(* IEC 61131-3 sources: plc-st-coding-agent/progress/evidence/f14_v2_public_20261112b/jobs/codex_minimax-m27, 5 files *)

(* ---- public-easy-01.candidate_01.st ---- *)
FUNCTION_BLOCK FillingLineControl
VAR_INPUT
    bottleSensor           : BOOL;
    cleaningConfirmButton  : BOOL;
    fillingConfirmButton   : BOOL;
    cappingConfirmButton   : BOOL;
    packingConfirmButton   : BOOL;
    finishedButton         : BOOL;
END_VAR

VAR_OUTPUT
    Pump_Motor     : BOOL := FALSE;
    Filling_Valve  : BOOL := FALSE;
    Capping_Machine: BOOL := FALSE;
    Packing_Machine: BOOL := FALSE;
    Completion_Light: BOOL := FALSE;
END_VAR

VAR
    state : INT := 0;
    lastBottleSensor : BOOL := FALSE;
END_VAR

    // Detect bottle arrival
    IF bottleSensor AND NOT lastBottleSensor THEN
        state := 1;
    END_IF
    lastBottleSensor := bottleSensor;

    // State machine
    CASE state OF
        0:  // IDLE
            Pump_Motor := FALSE;
            Filling_Valve := FALSE;
            Capping_Machine := FALSE;
            Packing_Machine := FALSE;
            Completion_Light := FALSE;

        1:  // CLEANING
            Pump_Motor := TRUE;
            Filling_Valve := FALSE;
            Capping_Machine := FALSE;
            Packing_Machine := FALSE;
            Completion_Light := FALSE;
            IF cleaningConfirmButton THEN
                state := 2;
            END_IF

        2:  // FILLING
            Pump_Motor := FALSE;
            Filling_Valve := TRUE;
            Capping_Machine := FALSE;
            Packing_Machine := FALSE;
            Completion_Light := FALSE;
            IF fillingConfirmButton THEN
                state := 3;
            END_IF

        3:  // CAPPING
            Pump_Motor := FALSE;
            Filling_Valve := FALSE;
            Capping_Machine := TRUE;
            Packing_Machine := FALSE;
            Completion_Light := FALSE;
            IF cappingConfirmButton THEN
                state := 4;
            END_IF

        4:  // PACKING
            Pump_Motor := FALSE;
            Filling_Valve := FALSE;
            Capping_Machine := FALSE;
            Packing_Machine := TRUE;
            Completion_Light := FALSE;
            IF packingConfirmButton THEN
                state := 5;
            END_IF

        5:  // COMPLETE
            Pump_Motor := FALSE;
            Filling_Valve := FALSE;
            Capping_Machine := FALSE;
            Packing_Machine := FALSE;
            Completion_Light := TRUE;
            IF finishedButton THEN
                state := 0;
            END_IF
    END_CASE
END_FUNCTION_BLOCK

(* ---- public-easy-01.candidate_02.st ---- *)
FUNCTION_BLOCK FillingLineControl
VAR_INPUT
    bottleSensor           : BOOL;
    cleaningConfirmButton  : BOOL;
    fillingConfirmButton   : BOOL;
    cappingConfirmButton   : BOOL;
    packingConfirmButton   : BOOL;
    finishedButton         : BOOL;
END_VAR

VAR_OUTPUT
    Pump_Motor      : BOOL := FALSE;
    Filling_Valve   : BOOL := FALSE;
    Capping_Machine : BOOL := FALSE;
    Packing_Machine : BOOL := FALSE;
    Completion_Light: BOOL := FALSE;
END_VAR

VAR
    state               : INT := 0;
    lastBottleSensor    : BOOL := FALSE;
    lastCleaningButton  : BOOL := FALSE;
    lastFillingButton   : BOOL := FALSE;
    lastCappingButton   : BOOL := FALSE;
    lastPackingButton   : BOOL := FALSE;
    lastFinishedButton  : BOOL := FALSE;
END_VAR

    // Detect bottle arrival on rising edge
    IF bottleSensor AND NOT lastBottleSensor THEN
        state := 1;
    END_IF
    lastBottleSensor := bottleSensor;

    // State machine
    CASE state OF
        0:  // IDLE
            Pump_Motor := FALSE;
            Filling_Valve := FALSE;
            Capping_Machine := FALSE;
            Packing_Machine := FALSE;
            Completion_Light := FALSE;

        1:  // CLEANING
            Pump_Motor := TRUE;
            Filling_Valve := FALSE;
            Capping_Machine := FALSE;
            Packing_Machine := FALSE;
            Completion_Light := FALSE;
            // Rising edge detection for button
            IF cleaningConfirmButton AND NOT lastCleaningButton THEN
                state := 2;
            END_IF

        2:  // FILLING
            Pump_Motor := FALSE;
            Filling_Valve := TRUE;
            Capping_Machine := FALSE;
            Packing_Machine := FALSE;
            Completion_Light := FALSE;
            // Rising edge detection for button
            IF fillingConfirmButton AND NOT lastFillingButton THEN
                state := 3;
            END_IF

        3:  // CAPPING
            Pump_Motor := FALSE;
            Filling_Valve := FALSE;
            Capping_Machine := TRUE;
            Packing_Machine := FALSE;
            Completion_Light := FALSE;
            // Rising edge detection for button
            IF cappingConfirmButton AND NOT lastCappingButton THEN
                state := 4;
            END_IF

        4:  // PACKING
            Pump_Motor := FALSE;
            Filling_Valve := FALSE;
            Capping_Machine := FALSE;
            Packing_Machine := TRUE;
            Completion_Light := FALSE;
            // Rising edge detection for button
            IF packingConfirmButton AND NOT lastPackingButton THEN
                state := 5;
            END_IF

        5:  // COMPLETE
            Pump_Motor := FALSE;
            Filling_Valve := FALSE;
            Capping_Machine := FALSE;
            Packing_Machine := FALSE;
            Completion_Light := TRUE;
            // Rising edge detection for button
            IF finishedButton AND NOT lastFinishedButton THEN
                state := 0;
            END_IF
    END_CASE

    // Update last button states for edge detection
    lastCleaningButton := cleaningConfirmButton;
    lastFillingButton := fillingConfirmButton;
    lastCappingButton := cappingConfirmButton;
    lastPackingButton := packingConfirmButton;
    lastFinishedButton := finishedButton;
END_FUNCTION_BLOCK

(* ---- public-easy-02.candidate_01.st ---- *)
FUNCTION_BLOCK FB_DualWordEdgeDetection
VAR_INPUT
    value : DWORD;
END_VAR

VAR_OUTPUT
    hasChanged      : BOOL;
    hasRisingEdges  : BOOL;
    risingBits      : DWORD;
    noOfRisingBits  : USINT;
    hasFallingEdges : BOOL;
    fallingBits     : DWORD;
    noOfFallingBits : USINT;
END_VAR

VAR
    prevValue    : DWORD;
    changedBits  : DWORD;
    bitPosition  : USINT;
    bitMask      : DWORD;
END_VAR

changedBits := value XOR prevValue;

risingBits  := changedBits AND value;
fallingBits := changedBits AND NOT value;

hasChanged      := (value <> prevValue);
hasRisingEdges  := (risingBits  <> 0);
hasFallingEdges := (fallingBits <> 0);

noOfRisingBits  := 0;
noOfFallingBits := 0;

FOR bitPosition := 0 TO 31 DO
    bitMask := SHL(DWORD#1, bitPosition);
    IF (risingBits AND bitMask) <> DWORD#0 THEN
        noOfRisingBits := noOfRisingBits + 1;
    END_IF
    IF (fallingBits AND bitMask) <> DWORD#0 THEN
        noOfFallingBits := noOfFallingBits + 1;
    END_IF
END_FOR

prevValue := value;

END_FUNCTION_BLOCK

(* ---- public-easy-03.candidate_01.st ---- *)
FUNCTION_BLOCK AlarmHysteresis
VAR_INPUT
    Value       : REAL;
    hiLevel     : REAL;
    loLevel     : REAL;
    hystWindow  : REAL;
END_VAR

VAR_OUTPUT
    hiAlarm     : BOOL;
    loAlarm     : BOOL;
    error       : BOOL;
    status      : WORD;
END_VAR

    // Error checking: loLevel must be less than hiLevel
    IF loLevel >= hiLevel THEN
        error := TRUE;
        status := 16#8001;
        RETURN;
    END_IF

    // Error checking: hystWindow must be less than the range between hiLevel and loLevel
    IF hystWindow >= (hiLevel - loLevel) THEN
        error := TRUE;
        status := 16#8002;
        RETURN;
    END_IF

    // No error
    error := FALSE;
    status := 16#0000;

    // High alarm logic with hysteresis
    // Trigger: Value > hiLevel
    // Release: Value < hiLevel - hystWindow
    IF Value > hiLevel THEN
        hiAlarm := TRUE;
    ELSIF Value < (hiLevel - hystWindow) THEN
        hiAlarm := FALSE;
    END_IF

    // Low alarm logic with hysteresis
    // Trigger: Value < loLevel
    // Release: Value > loLevel + hystWindow
    IF Value < loLevel THEN
        loAlarm := TRUE;
    ELSIF Value > (loLevel + hystWindow) THEN
        loAlarm := FALSE;
    END_IF

END_FUNCTION_BLOCK

(* ---- public-easy-03.candidate_02.st ---- *)
FUNCTION_BLOCK AlarmHysteresis
VAR_INPUT
    Value       : REAL;
    hiLevel     : REAL;
    loLevel     : REAL;
    hystWindow  : REAL;
END_VAR

VAR_OUTPUT
    hiAlarm     : BOOL := FALSE;
    loAlarm     : BOOL := FALSE;
    error       : BOOL;
    status      : WORD := 16#0000;
END_VAR

    // Error: loLevel must be less than hiLevel
    IF loLevel >= hiLevel THEN
        error := TRUE;
        status := 16#8001;
        RETURN;
    END_IF

    // Error: hystWindow must be less than the deviation range
    IF hystWindow >= (hiLevel - loLevel) THEN
        error := TRUE;
        status := 16#8002;
        RETURN;
    END_IF

    // No error - only clear error flag, preserve status
    error := FALSE;

    // High alarm with hysteresis
    // Trigger: Value > hiLevel
    // Release: Value < hiLevel - hystWindow
    IF Value > hiLevel THEN
        hiAlarm := TRUE;
    ELSIF Value < (hiLevel - hystWindow) THEN
        hiAlarm := FALSE;
    END_IF

    // Low alarm with hysteresis
    // Trigger: Value < loLevel
    // Release: Value > loLevel + hystWindow
    IF Value < loLevel THEN
        loAlarm := TRUE;
    ELSIF Value > (loLevel + hystWindow) THEN
        loAlarm := FALSE;
    END_IF

END_FUNCTION_BLOCK
